(* IEC 61131-3 sources: codesys-framework/txt/application/WeVe General (library)/Blink/FB_BlinkService, 1 file *)

(* ---- Blinks.prop.st ---- *)
PROPERTY Blinks : SC_Blinks

// --- BEGIN IMPLEMENTATION ---

// ----------- GET -----------
VAR
END_VAR

// -- BEGIN IMPLEMENTATION GET --
Blinks := _scBlinks;
